FUNCTION_BLOCK FakeClock IMPLEMENTS I_Clock
VAR
    _Now : LTIME;
END_VAR
(*
    FakeClock

    Stands still until the test moves it.
*)

METHOD PUBLIC Advance
VAR_INPUT
    Duration : LTIME;
END_VAR
_Now := _Now + Duration;
END_METHOD

PROPERTY PUBLIC Now : LTIME
GET
Now := _Now;
END_GET
END_PROPERTY

END_FUNCTION_BLOCK

(* stored: Version 1.1.0.1, ProductVersion 3.1.4026.0
   POU FakeClock: Id {dbeb2fd8-2ceb-4323-8f60-c29685dc72ca}, SpecialFunc None
   Folder I_Clock: Id {ea1665d9-4a76-4cb0-a728-2a6225e5e28e}
   Method Advance: Id {d9debce1-9baf-4e9c-999e-cf2dc60fd16d}
   Property Now: Id {770be202-787b-425e-8f10-82f6dd7ba35b}
   Get Get: Id {7745eb38-7646-4093-b4ce-16f51637c250} *)
